(* IEC 61131-3 sources: llm-plc-st-eval/data/sonda_gemini/gemini-3.1-pro-preview/A6/zero_shot, 3 files *)

(* ---- ejec_1.st ---- *)
```iecst
FUNCTION_BLOCK FB_Modos
VAR_INPUT
    selector : INT;
    estadoSeguro : BOOL;
    cmdAuto : ARRAY[0..7] OF BOOL;
    cmdManual : ARRAY[0..7] OF BOOL;
    idxForzado : INT;
    valorForzado : BOOL;
    confirmarForzado : BOOL;
END_VAR

VAR_OUTPUT
    modoActivo : INT := 1; // Inicializa en modo manual (1) por defecto
    actuador : ARRAY[0..7] OF BOOL;
END_VAR

VAR
    prevConfirmar : BOOL;
    flancoConfirmar : BOOL;
    prevModo : INT := 1;
    i : INT;
END_VAR

// Detección de flanco de subida para la señal de confirmación de forzado
flancoConfirmar := confirmarForzado AND NOT prevConfirmar;
prevConfirmar := confirmarForzado;

// Gestión de cambio de modo de operación (solo si hay estado seguro y el selector es válido)
IF estadoSeguro THEN
    IF (selector >= 0) AND (selector <= 2) THEN
        modoActivo := selector;
    END_IF;
END_IF;

// Lógica de control de actuadores según el modo activo
CASE modoActivo OF
    0: // Modo Automático
        FOR i := 0 TO 7 DO
            actuador[i] := cmdAuto[i];
        END_FOR;

    1: // Modo Manual
        FOR i := 0 TO 7 DO
            actuador[i] := cmdManual[i];
        END_FOR;

    2: // Modo Mantenimiento
        // Al entrar al modo mantenimiento, todos los actuadores parten apagados
        IF prevModo <> 2 THEN
            FOR i := 0 TO 7 DO
                actuador[i] := FALSE;
            END_FOR;
        END_IF;

        // Si se pierde el estado seguro durante el mantenimiento, se anulan los forzados
        IF NOT estadoSeguro THEN
            FOR i := 0 TO 7 DO
                actuador[i] := FALSE;
            END_FOR;
        ELSE
            // Aplicar forzado individual en flanco de subida si el índice está en rango
            IF flancoConfirmar THEN
                IF (idxForzado >= 0) AND (idxForzado <= 7) THEN
                    actuador[idxForzado] := valorForzado;
                END_IF;
            END_IF;
        END_IF;
END_CASE;

// Actualizar el registro del modo previo para evaluar transiciones en el siguiente ciclo
prevModo := modoActivo;

END_FUNCTION_BLOCK
```

(* ---- ejec_2.st ---- *)
```iecst
FUNCTION_BLOCK FB_Modos
VAR_INPUT
    selector : INT; (* 0: Auto, 1: Manual, 2: Mantenimiento *)
    estadoSeguro : BOOL; (* Condición para permitir cambio de modo *)
    cmdAuto : ARRAY[0..7] OF BOOL; (* Comandos en modo automático *)
    cmdManual : ARRAY[0..7] OF BOOL; (* Comandos en modo manual *)
    idxForzado : INT; (* Índice del actuador a forzar (0-7) *)
    valorForzado : BOOL; (* Valor a aplicar al actuador forzado *)
    confirmarForzado : BOOL; (* Señal para aplicar el forzado *)
END_VAR

VAR_OUTPUT
    modoActivo : INT := 1; (* Modo vigente, inicializado en Manual (1) *)
    actuador : ARRAY[0..7] OF BOOL; (* Estado de los 8 actuadores *)
END_VAR

VAR
    trigConfirmar : R_TRIG; (* Detector de flanco de subida para confirmarForzado *)
    modoAnterior : INT := 1; (* Memoria del modo en el ciclo anterior *)
    i : INT; (* Variable para bucles *)
END_VAR

(* 1. Gestión del cambio de modo de operación *)
IF estadoSeguro THEN
    IF selector >= 0 AND selector <= 2 THEN
        modoActivo := selector;
    END_IF;
END_IF;

(* 2. Detección de flanco para la confirmación de forzado *)
trigConfirmar(CLK := confirmarForzado);

(* 3. Lógica de control de actuadores según el modo activo *)
CASE modoActivo OF

    0: (* MODO AUTOMÁTICO *)
        FOR i := 0 TO 7 DO
            actuador[i] := cmdAuto[i];
        END_FOR;

    1: (* MODO MANUAL *)
        FOR i := 0 TO 7 DO
            actuador[i] := cmdManual[i];
        END_FOR;

    2: (* MODO MANTENIMIENTO *)
        (* Al entrar al modo mantenimiento, apagar todos los actuadores *)
        IF modoAnterior <> 2 THEN
            FOR i := 0 TO 7 DO
                actuador[i] := FALSE;
            END_FOR;
        END_IF;

        (* Si se pierde el estado seguro, anular forzados y apagar actuadores *)
        IF NOT estadoSeguro THEN
            FOR i := 0 TO 7 DO
                actuador[i] := FALSE;
            END_FOR;
        ELSE
            (* Aplicar forzado individual en flanco de subida si el índice es válido *)
            IF trigConfirmar.Q THEN
                IF idxForzado >= 0 AND idxForzado <= 7 THEN
                    actuador[idxForzado] := valorForzado;
                END_IF;
            END_IF;
        END_IF;

END_CASE;

(* 4. Actualización de la memoria del modo para el próximo ciclo *)
(* Nota: Al salir de mantenimiento (modoActivo pasa a 0 o 1), los forzados se anulan
   automáticamente al sobrescribirse el array actuador con cmdAuto o cmdManual *)
modoAnterior := modoActivo;

END_FUNCTION_BLOCK
```

(* ---- ejec_3.st ---- *)
```iecst
FUNCTION_BLOCK FB_Modos
VAR_INPUT
    selector : INT;
    estadoSeguro : BOOL;
    cmdAuto : ARRAY[0..7] OF BOOL;
    cmdManual : ARRAY[0..7] OF BOOL;
    idxForzado : INT;
    valorForzado : BOOL;
    confirmarForzado : BOOL;
END_VAR

VAR_OUTPUT
    modoActivo : INT := 1; // El modo vigente al arrancar es manual (1)
    actuador : ARRAY[0..7] OF BOOL;
END_VAR

VAR
    i : INT;
    modoAnterior : INT := 1;
    prevConfirmar : BOOL := FALSE;
    flancoConfirmar : BOOL;
END_VAR

// 1. Gestión de cambio de modo de operación
IF estadoSeguro THEN
    // Solo se aceptan valores válidos (0=Auto, 1=Manual, 2=Mantenimiento)
    IF selector >= 0 AND selector <= 2 THEN
        modoActivo := selector;
    END_IF;
END_IF;

// 2. Detección de flanco de subida para la señal de confirmación
flancoConfirmar := confirmarForzado AND NOT prevConfirmar;
prevConfirmar := confirmarForzado;

// 3. Inicialización al entrar en modo mantenimiento (apagar todos)
IF modoActivo = 2 AND modoAnterior <> 2 THEN
    FOR i := 0 TO 7 DO
        actuador[i] := FALSE;
    END_FOR;
END_IF;

// 4. Lógica de control de actuadores según el modo activo
CASE modoActivo OF
    0: // Modo Automático
        FOR i := 0 TO 7 DO
            actuador[i] := cmdAuto[i];
        END_FOR;

    1: // Modo Manual
        FOR i := 0 TO 7 DO
            actuador[i] := cmdManual[i];
        END_FOR;

    2: // Modo Mantenimiento
        IF NOT estadoSeguro THEN
            // Si se pierde el estado seguro durante el mantenimiento, apagar todo
            FOR i := 0 TO 7 DO
                actuador[i] := FALSE;
            END_FOR;
        ELSE
            // Si hay flanco de subida y el índice está en rango, aplicar forzado
            IF flancoConfirmar THEN
                IF idxForzado >= 0 AND idxForzado <= 7 THEN
                    actuador[idxForzado] := valorForzado;
                END_IF;
            END_IF;
        END_IF;
END_CASE;

// 5. Actualizar el modo anterior para el siguiente ciclo de escaneo
modoAnterior := modoActivo;

END_FUNCTION_BLOCK
```
